(* IEC 61131-3 sources: iolistgen/tests_support/pl_stub/src/DUTs/Motor, 6 files *)

(* ---- E_MotorAlarm.dut.st ---- *)
// Назначение: заглушка plc-process-lib 1.0.0 для проверки типов сгенерированного кода без CODESYS
//             (API.md, раздел 4.1); не библиотека — тел и внутренних переменных нет
// Автор:      kr0nsch
// Версия:     1.0.0 (выпуск библиотеки)
// Документ:   docs/GENERATORS.md, раздел «Проверка ST без CODESYS»
{attribute 'qualified_only'}
TYPE E_MotorAlarm :
(
    FailToStart := 0,
    FeedbackLost := 1,
    FailToStop := 2,
    UncommandedRun := 3,
    ExtFault := 4,
    InterlockTrip := 5,
    CommLoss := 6,
    SpeedDeviation := 7
) UINT;
END_TYPE

(* ---- E_MotorState.dut.st ---- *)
// Назначение: заглушка plc-process-lib 1.0.0 для проверки типов сгенерированного кода без CODESYS
//             (API.md, раздел 13.1); не библиотека — тел и внутренних переменных нет
// Автор:      kr0nsch
// Версия:     1.0.0 (выпуск библиотеки)
// Документ:   docs/GENERATORS.md, раздел «Проверка ST без CODESYS»
{attribute 'qualified_only'}
{attribute 'strict'}
TYPE E_MotorState :
(
    Stopped := 0,
    Starting := 1,
    Running := 2,
    Stopping := 3,
    Fault := 4
) INT;
END_TYPE

(* ---- ST_MotorCfg.dut.st ---- *)
// Назначение: заглушка plc-process-lib 1.0.0 для проверки типов сгенерированного кода без CODESYS
//             (API.md, раздел 13.1); не библиотека — тел и внутренних переменных нет
// Автор:      kr0nsch
// Версия:     1.0.0 (выпуск библиотеки)
// Документ:   docs/GENERATORS.md, раздел «Проверка ST без CODESYS»
{attribute 'qualified_only'}
TYPE ST_MotorCfg :
STRUCT
    xFbUsed            : BOOL := TRUE;
    tFbStart           : TIME := T#5S;
    tFbStop            : TIME := T#5S;
    tFbLossFilter      : TIME := T#500MS;
    tExtFaultFilter    : TIME := T#200MS;
    tMinRun            : TIME := T#0S;
    tMinStop           : TIME := T#0S;
    uiMaxStartsPerHour : UINT := 0;
    tResetWindow       : TIME := T#3S;
    tResetPulse        : TIME := T#1S;
    wInterlockMask     : WORD := 16#FFFF;
    wPermitMask        : WORD := 16#FFFF;
    udiMaintInterval_h : UDINT := 0;
    udiMaintStarts     : UDINT := 0;
    stVfd              : ST_VfdCfg;
    udiAlarmIdBase     : UDINT := 0;
    // lint:allow STL007 имя массива по контракту API.md (префикс a + тип элемента)
    astAlarm       : ARRAY[0..GVL_Const.DEV_ALARMS_MAX - 1] OF ST_AlarmCfg := [
            (ePriority := E_AlarmPriority.Medium),
            (ePriority := E_AlarmPriority.Medium),
            (ePriority := E_AlarmPriority.High),
            (ePriority := E_AlarmPriority.High),
            (ePriority := E_AlarmPriority.Medium),
            (ePriority := E_AlarmPriority.None),
            (ePriority := E_AlarmPriority.Medium),
            (ePriority := E_AlarmPriority.Low)];
END_STRUCT
END_TYPE

(* ---- ST_MotorCmd.dut.st ---- *)
// Назначение: заглушка plc-process-lib 1.0.0 для проверки типов сгенерированного кода без CODESYS
//             (API.md, раздел 13.1); не библиотека — тел и внутренних переменных нет
// Автор:      kr0nsch
// Версия:     1.0.0 (выпуск библиотеки)
// Документ:   docs/GENERATORS.md, раздел «Проверка ST без CODESYS»
{attribute 'qualified_only'}
TYPE ST_MotorCmd :
STRUCT
    stCommon     : ST_DeviceCmd;
    xStart       : BOOL;
    xStop        : BOOL;
    xResetMaint  : BOOL;
    rSpeedSp_pct : REAL;
END_STRUCT
END_TYPE

(* ---- ST_MotorSts.dut.st ---- *)
// Назначение: заглушка plc-process-lib 1.0.0 для проверки типов сгенерированного кода без CODESYS
//             (API.md, раздел 13.1); не библиотека — тел и внутренних переменных нет
// Автор:      kr0nsch
// Версия:     1.0.0 (выпуск библиотеки)
// Документ:   docs/GENERATORS.md, раздел «Проверка ST без CODESYS»
{attribute 'qualified_only'}
TYPE ST_MotorSts :
STRUCT
    stCommon          : ST_DeviceSts;
    eState            : E_MotorState;
    wInterlock        : WORD;
    wPermitMissing    : WORD;
    uiFirstOut        : UINT;
    uiInhibitRemain_s : UINT;
    uiStartsLastHour  : UINT;
    rRunTime_h        : REAL;
    udiStarts         : UDINT;
    rRunTimeMaint_h   : REAL;
    udiStartsMaint    : UDINT;
    rSpeedRef_pct     : REAL;
    rSpeedAct_pct     : REAL;
    udiRunCurrent_s   : UDINT;
END_STRUCT
END_TYPE

(* ---- ST_VfdCfg.dut.st ---- *)
// Назначение: заглушка plc-process-lib 1.0.0 для проверки типов сгенерированного кода без CODESYS
//             (API.md, раздел 13.1); не библиотека — тел и внутренних переменных нет
// Автор:      kr0nsch
// Версия:     1.0.0 (выпуск библиотеки)
// Документ:   docs/GENERATORS.md, раздел «Проверка ST без CODESYS»
{attribute 'qualified_only'}
TYPE ST_VfdCfg :
STRUCT
    rSpeedMin_pct    : REAL := 0.0;
    rSpeedMax_pct    : REAL := 100.0;
    rRampUp_pctps    : REAL := 0.0;
    rRampDown_pctps  : REAL := 0.0;
    xFbFromComm      : BOOL := TRUE;
    xCommLossIsFault : BOOL := TRUE;
    tCommLoss        : TIME := T#3S;
    rSpeedDev_pct    : REAL := 10.0;
    tSpeedDev        : TIME := T#10S;
END_STRUCT
END_TYPE
